                          CallSubProgram
                          PROCESS_Step := 0
                          WRK_Done := True
                    Case (caseValue=20)
                      SuppressedNode
                        Folder Biorad rack
                          'load racks'
                          If Task_ID≟16
                            SuppressedNode
                              PRC_RackCounter := 0
                            Loop While (checkContinuously=false) expression=(PRC_RackCounter<PRC_RackNumber) and  not CMD_Stop
                              JIG_Slot := PRC_RackCounter
                              Action := 1
                              PRC_Target := 0
                              CallSubProgram
                              If OBJ_Picked
                                Action := 2
                                PRC_Target := 1
                                CallSubProgram
                                Action := 7
                                PRC_Target := 1
                                CallSubProgram
                                PRC_RackCounter := PRC_RackCounter+1
                            WRK_Done := True
                            PROCESS_Step := 0
                          'unload racks'
                          SuppressedNode
                            If Task_ID≟17
                              SuppressedNode
                                PRC_RackCounter := 0
                              Loop While (checkContinuously=false) expression=(PRC_RackCounter<PRC_RackNumber) and  not CMD_Stop
                                JIG_Slot := PRC_RackCounter
                                Action := 8
                                PRC_Target := 1
                                Script: textmsg("Callactionunload=",Action)
                                CallSubProgram
                                Action := 1
                                PRC_Target := 1
                                Script: textmsg("Callactionpick=",Action)
                                CallSubProgram
                                If OBJ_Picked
                                  Action := 2
                                  PRC_Target := 0
                                  Script: textmsg("Callactionplace=",Action)
                                  CallSubProgram
                                  PRC_RackCounter := PRC_RackCounter+1
                              WRK_Done := True
                              PROCESS_Step := 0
                          If Task_ID≟17
                            PRC_RackCounter := 0
                            Loop While (checkContinuously=false) expression=(PRC_RackCounter<PRC_RackNumber) and  not CMD_Stop
                              Wait Condition expression=SensorData[PRC_RackCounter]≟1
                              JIG_Slot := PRC_RackCounter
                              Action := 8
                              PRC_Target := 1
                              Script: textmsg("Callactionunload=",Action)
                              CallSubProgram
                              Action := 1
                              PRC_Target := 1
                              Script: textmsg("Callactionpick=",Action)
                              CallSubProgram
                              If OBJ_Picked
                                Action := 2
                                PRC_Target := 0
                                Script: textmsg("Callactionplace=",Action)
                                CallSubProgram
                                PRC_RackCounter := PRC_RackCounter+1
                            WRK_Done := True
                            PROCESS_Step := 0
                    Case (caseValue=43)
                      SuppressedNode
                        Folder Pick the rack
                          Action := 131
                          CallSubProgram
                          Action := 1
                          CallSubProgram
                          PROCESS_Step := 0
                          WRK_Done := True
                    Case (caseValue=2147483647)
                      WRK_Done := True
                      PROCESS_Step := 0
          If CMD_Hold
            STATE := 9
            Script: ugo_update_outputs()
          ElseIf CMD_Suspend
            STATE := 12
            Script: ugo_update_outputs()
      Case (caseValue=7)
        Folder Completing [hidden by the author, left out]
      Case (caseValue=8)
        Folder Complete [hidden by the author, left out]
      Case (caseValue=9)
        Folder Holding [hidden by the author, left out]
      Case (caseValue=10)
        Folder Held [hidden by the author, left out]
      Case (caseValue=11)
        Folder Unholding [hidden by the author, left out]
      Case (caseValue=12)
        Folder Suspending [hidden by the author, left out]
      Case (caseValue=13)
        Folder Suspended [hidden by the author, left out]
      Case (caseValue=14)
        Folder Unsuspending [hidden by the author, left out]
      Case (caseValue=15)
        Folder Aborting [hidden by the author, left out]
      Case (caseValue=16)
        Folder Aborted [hidden by the author, left out]
      Case (caseValue=17)
        Folder Clearing [hidden by the author, left out]
    Script: log_state(STATE_Info)
    Script: log_warning(WARNING.MSG)
    Script: log_error(ERROR.MSG)
    Folder Times [hidden by the author, left out]
    SuppressedNode
      Script: sync()
    Wait Sleep waitTime=0.1
Thread Thread_1 (runOnlyOnce=false)
  Folder Dosing Weight
    If Start_thread≟ True
      weight_value := get_weight()
      diff := target_weight-weight_value
      Wait Sleep waitTime=0.2
      Script: sync()
  Script: sync()
Thread Thread_2 (runOnlyOnce=false)
  Folder Vibration motor
    Loop While (checkContinuously=true) expression=vib_thread≟ True
      diff := target_weight-weight_value
      If diff>0.02 and spatula≠"spatula_flat_S" (checkContinuously=true)
        SuppressedNode
          Script: vibration_4()
        Set AnalogOutput pin=analog_out[0]; analogValue=4
      ElseIf diff>0.02 and spatula≟"spatula_flat_S"
        Script: vibration_3()
      ElseIf diff≤0.03 (checkContinuously=true)
        Script: vibration_2()
      Else 
        Set AnalogOutput pin=analog_out[0]; analogValue=0
  Script: sync()
Thread Thread_3 (runOnlyOnce=false)
  Folder Container weight
    If w_full_thread≟ True
      aa_weight_cont := get_cont_weight()
      Wait Sleep waitTime=0.2
      Script: sync()
  Script: sync()
SubProgram  [hidden by the author, left out]
SubProgram  [hidden by the author, left out]
SubProgram -> Sub_Action_V4
